Fanuc KAREL source: KT00751.KL

PROGRAM KT00751
%NOLOCKGROUP
VAR
  R1: REAL
  R2: REAL
  OUT: REAL
BEGIN
  R1 = 2.0
  R2 = 3.0
  R1 = 2.0
  R2 = 3.0
  OUT = ABS(R1)
END KT00751
